FUNCTION FC 1 : VOID
BEGIN
      A I 0.0
END_FUNCTION
